(* IEC 61131-3 sources: soft_bellows/soft_bellows_plc/Temp/History/Logical/05_23_2024_10_09_03/basic_pneu_stand/Riadenie/Program, 4 files *)

(* ---- Cyclic.st ---- *)
PROGRAM _CYCLIC

	IF tlacidla.zapni=TRUE THEN

		FOR i:=0 TO 7 BY 1 DO
			regulatory.reg[i] := REAL_TO_INT(display.in_reg[i]/100*32765/9);
		END_FOR

	ELSE

		FOR i:=0 TO 3 BY 1 DO
			tlacidla.ventil[i] := FALSE;
		END_FOR

		FOR i:=0 TO 7 BY 1 DO
			regulatory.reg[i] := 0;
		END_FOR

	END_IF

END_PROGRAM

(* ---- Exit.st ---- *)
PROGRAM _EXIT
	(* Insert code here *)

END_PROGRAM

(* ---- Init.st ---- *)
PROGRAM _INIT
	(* Insert code here *)

END_PROGRAM

(* ---- Variables.var ---- *)
VAR
	i : INT;
END_VAR
